TYPE ST_EL6910HistoryRow :
STRUCT
    sSeverity : STRING(16);
    sTimestamp : STRING(32);
    sMessage : STRING(255);
    sDetail : STRING(255);
END_STRUCT
END_TYPE

(* stored: Version 1.1.0.1, ProductVersion 3.1.4026.18
   DUT ST_EL6910HistoryRow: Id {ac93aed0-1c5a-431a-a899-e746be378fae} *)
